(*
SPDX-FileCopyrightText: © 2026 Oleksandr Tiutyk <trofimich@gmail.com>
SPDX-License-Identifier: MIT
License: https://opensource.org/license/mit
*)

(*!
<summary>Provides controlled execution and formatter failures for workflow contract tests.</summary>
<description>
Persistent test instances own their borrowed configuration and exception template. No hardware effects or
terminal allocation injection are performed. The fixture can defer its initial resetting step. All observations are task-local.
</description>
*)

{attribute 'enable_dynamic_creation'}
{attribute 'no_explicit_call' := 'do not call this function block directly'}
{attribute 'no_assign'}
FUNCTION_BLOCK WorkflowContractActivity EXTENDS TOF_Workflow.Activity
VAR_INPUT
	//! <summary>Raises an ordinary work exception on every running call while enabled.</summary>
	throwOrdinaryFailure : BOOL;
	//! <summary>Raises a concrete exception whose message formatter itself raises.</summary>
	throwMessageFailure : BOOL;
	//! <summary>Completes running immediately when no injected failure is enabled.</summary>
	completeRunning : BOOL;
	//! <summary>Keeps the first reset step pending until the next Execute call.</summary>
	deferFirstResetStep : BOOL;
	//! <summary>Optional persistent observer incremented on ordinary destruction of a factory fixture.</summary>
	exitCount : REFERENCE TO DINT;
END_VAR
VAR_OUTPUT
	//! <summary>Number of fresh or resumed start callbacks.</summary>
	startCount : DINT;
	//! <summary>Number of running callbacks, including entry calls.</summary>
	runningCount : DINT;
	//! <summary>Number of stopping callbacks.</summary>
	stopCount : DINT;
END_VAR
VAR_STAT
	//! <summary>Initialized static metadata available during inherited base initialization.</summary>
	_ClassName : STRING := __POUNAME();
END_VAR
VAR
	_MessageFailure : ThrowingGetMessageException;
END_VAR

(*!
<summary>Returns the initialized static name of this concrete fixture.</summary>
*)
{attribute 'monitoring' := 'call'}
PROPERTY ClassName : REFERENCE TO STRING
GET
ClassName REF= _ClassName;
END_GET
END_PROPERTY

(*!
<summary>Borrows the test project namespace without changing it.</summary>
*)
{attribute 'monitoring' := 'call'}
PROPERTY NamespaceName : REFERENCE TO STRING
GET
NamespaceName REF= CurrentNamespace.Name;
END_GET
END_PROPERTY

(*!
<summary>Reports the size of this concrete fixture in bytes.</summary>
*)
{attribute 'monitoring' := 'call'}
PROPERTY SelfSize : ULINT
GET
SelfSize := XSIZEOF(THIS^);
END_GET
END_PROPERTY

(*!
<summary>Counts execution and produces the selected ordinary result or exception.</summary>
<param name="startRunning">Marks a fresh start for the entry counter.</param>
<param name="startResuming">Marks a resumed start for the entry counter.</param>
<param name="haltReason">Unused because this probe does not halt.</param>
*)
METHOD PROTECTED OnRunning : TOF_Workflow.ACTIVITY_RUNNING_STATE
VAR_INPUT
	startRunning : BOOL;
	startResuming : BOOL;
END_VAR
VAR_OUTPUT
	haltReason : WSTRING(255);
END_VAR
runningCount := runningCount + 1;

IF startRunning OR_ELSE startResuming THEN
	startCount := startCount + 1;
END_IF

IF throwMessageFailure THEN
	_MessageFailure.Throw(
		sourceNamespaceName := NamespaceName,
		sourceClassName := ClassName,
		sourcePOUName := __POUNAME(),
		sourcePosition := __POSITION(),
		message := "Controlled original workflow failure"
	);
END_IF

IF throwOrdinaryFailure THEN
	TOF_Core.Exceptions.ThrowStandard(
		sourceNamespaceName := NamespaceName,
		sourceClassName := ClassName,
		sourcePOUName := __POUNAME(),
		sourcePosition := __POSITION(),
		message := "Controlled workflow work failure"
	);
END_IF

IF completeRunning THEN
	OnRunning := TOF_Workflow.ACTIVITY_RUNNING_STATE.WORK_COMPLETED;
END_IF
END_METHOD

(*!
<summary>Counts a cooperative stopping step and finishes it immediately.</summary>
<param name="startCancelling">Unused cancellation-entry marker; stopping is immediate.</param>
<param name="startSuspending">Unused suspension-entry marker; stopping is immediate.</param>
<param name="haltReason">Unused because this probe does not halt.</param>
*)
METHOD PROTECTED OnStopping : TOF_Workflow.ACTIVITY_STOPPING_STATE
VAR_INPUT
	startCancelling : BOOL;
	startSuspending : BOOL;
END_VAR
VAR_OUTPUT
	haltReason : WSTRING(255);
END_VAR
stopCount := stopCount + 1;

OnStopping := TOF_Workflow.ACTIVITY_STOPPING_STATE.WORK_STOPPED;
END_METHOD

(*!
<summary>Optionally defers reset completion by one step.</summary>
<param name="startResetting">TRUE only on entry to reset.</param>
*)
METHOD PROTECTED OnResetting : TOF_Workflow.ACTIVITY_RESETTING_STATE
VAR_INPUT
	startResetting : BOOL;
END_VAR
IF startResetting AND_THEN deferFirstResetStep THEN
	OnResetting := TOF_Workflow.ACTIVITY_RESETTING_STATE.WORK_IN_PROGRESS;
ELSE
	OnResetting := TOF_Workflow.ACTIVITY_RESETTING_STATE.WORK_RESET;
END_IF
END_METHOD

(*!
<summary>Reports ordinary destruction to an optional persistent counter.</summary>
<description>The suite keeps the counter alive until disposal. Counting a callback does not certify physical deallocation.</description>
<param name="bInCopyCode">TwinCAT online-change indicator.</param>
*)
METHOD FB_exit : BOOL
VAR_INPUT
	bInCopyCode : BOOL;
END_VAR
IF NOT bInCopyCode AND_THEN __ISVALIDREF(exitCount) THEN
	exitCount := exitCount + 1;
END_IF
END_METHOD

END_FUNCTION_BLOCK

(* stored: Version 1.1.0.1
   POU WorkflowContractActivity: Id {fc48c35f-b3fe-48fc-a3b8-9fa46130ab61}, SpecialFunc None
   Property ClassName: Id {f324e79c-1990-48c9-baa5-591f4b13816e}
   Get Get: Id {c772a3d1-61fa-48f7-8e2d-80699270d09e}
   Property NamespaceName: Id {1316c653-00dc-4db5-a8d4-854599c3b4db}
   Get Get: Id {ebf46ea7-60ac-4aca-a424-bf25c22d5a7b}
   Property SelfSize: Id {1ecd69e7-5167-4854-9308-7818ee34a490}
   Get Get: Id {fcb80205-decd-46c4-9d6a-69cdf69f1579}
   Method OnRunning: Id {b0d50bd3-956d-412d-91cd-614ac6032d67}
   Method OnStopping: Id {4142d322-abe0-496d-8c39-359c8a0bb792}
   Method OnResetting: Id {d907286b-3240-4df7-a2de-d2d9d9e0e7a4}
   Method FB_exit: Id {7310ebf6-2f69-4010-bbc9-8e626f7df266} *)
